(* IEC 61131-3 sources: codesys-framework/txt/application/ToDo/Utils/Moving Average/DUT, 1 file *)

(* ---- SC_SystemParametersMovingAverage.dut.st ---- *)
TYPE SC_SystemParametersMovingAverage :
STRUCT
	iNbrOfItemsForAverage 	: UINT;
END_STRUCT
END_TYPE
